TYPE "ST_AccessPolicy"
VERSION : 0.1
   STRUCT
      "Required" : Array[0..11] of DInt;
      "SessionTimeout" : Time := T#0ms;
   END_STRUCT;
END_TYPE
